(* IEC 61131-3 sources: llm-plc-st-eval/data/processed_definitivo/qwen2.5-coder_14b/B6/few_shot, 3 files *)

(* ---- ejec_1.st ---- *)
FUNCTION_BLOCK FB_Baliza
VAR_INPUT
    alarma : BOOL; (* Condicion de alarma *)
END_VAR
VAR_OUTPUT
    lampara : BOOL; (* Lámpara de la baliza *)
END_VAR
VAR
    tParpadeo : TP; (* Temporizador para el parpadeo *)
    estado : BOOL; (* Estado actual de la lámpara *)
END_VAR

(* Inicialización del temporizador *)
IF alarma THEN
    tParpadeo(IN := TRUE, PT := T#1S);
    estado := tParpadeo.Q;
    lampara := estado;
ELSE
    lampara := FALSE;
END_IF;
END_FUNCTION_BLOCK

(* ---- ejec_2.st ---- *)
FUNCTION_BLOCK FB_Baliza
VAR_INPUT
    alarma : BOOL; (* Condición de alarma *)
END_VAR
VAR_OUTPUT
    lampara : BOOL; (* Lámpara de la baliza *)
END_VAR
VAR
    tParpadeo : TP; (* Temporizador para el parpadeo *)
    estado : BOOL; (* Estado actual de la lámpara *)
END_VAR

(* Inicialización del temporizador *)
IF alarma THEN
    tParpadeo(IN := TRUE, PT := T#1S);
    estado := NOT estado; (* Cambia el estado de la lámpara *)
ELSE
    tParpadeo(IN := FALSE);
    estado := FALSE; (* Apaga la lámpara *)
END_IF;

(* Asigna el estado de la lámpara *)
lampara := estado AND alarma;
END_FUNCTION_BLOCK

(* ---- ejec_3.st ---- *)
FUNCTION_BLOCK FB_Baliza
VAR_INPUT
    alarma : BOOL; (* Condición de alarma *)
END_VAR
VAR_OUTPUT
    lampara : BOOL; (* Lámpara de la baliza *)
END_VAR
VAR
    tParpadeo : TP; (* Temporizador para el parpadeo *)
    estado : BOOL; (* Estado actual de la lámpara *)
END_VAR

(* Inicialización del temporizador *)
IF alarma THEN
    tParpadeo(IN := TRUE, PT := T#1S);
    estado := tParpadeo.Q;
    lampara := estado;
ELSE
    lampara := FALSE;
END_IF
END_FUNCTION_BLOCK
